FUNCTION_BLOCK LevelSensors (* Composite Function Block Type *)
  (* Standard: 61499-2 *)
  (* Version 0.0, 6/20/2016, Andrei, nxtControl GmbH, template *)
  PACKAGE Main;
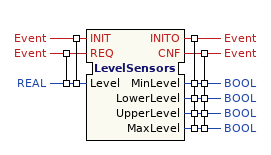
  EVENT_INPUT
    INIT WITH Level; (* Initialization Request *)
    REQ WITH Level; (* Normal Execution Request *)
  END_EVENT
  EVENT_OUTPUT
    INITO WITH MinLevel, LowerLevel, UpperLevel, MaxLevel; (* Initialization Confirm *)
    CNF WITH MinLevel, LowerLevel, UpperLevel, MaxLevel; (* Execution Confirmation *)
  END_EVENT
  VAR_INPUT
    Level : REAL; (* Input event qualifier *)
  END_VAR
  VAR_OUTPUT
    MinLevel : BOOL; (* Output event qualifier *)
    LowerLevel : BOOL;
    UpperLevel : BOOL;
    MaxLevel : BOOL;
  END_VAR
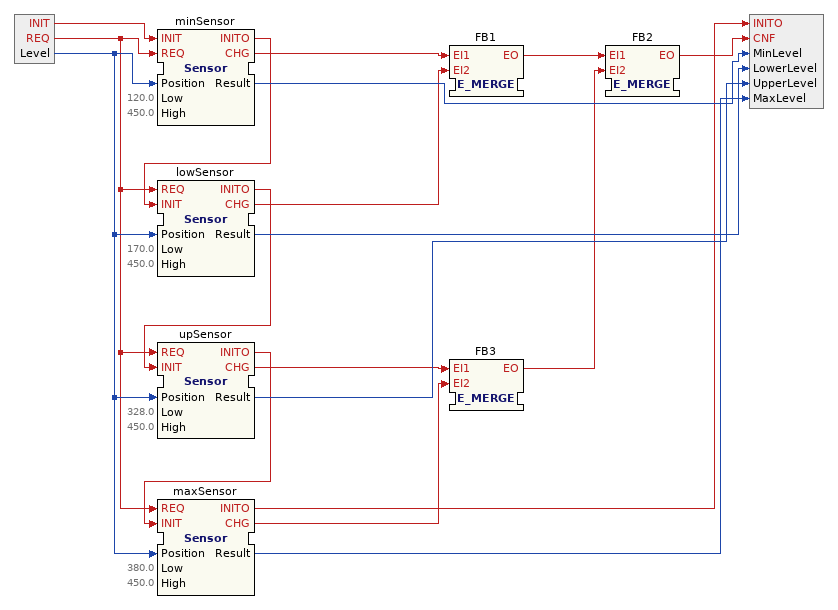
  FBS
    FB1 : E_MERGE;
    FB2 : E_MERGE;
    FB3 : E_MERGE;
    minSensor : Sensor(Low := 120.0, High := 450.0);
    lowSensor : Sensor(Low := 170.0, High := 450.0);
    upSensor : Sensor(Low := 328.0, High := 450.0);
    maxSensor : Sensor(Low := 380.0, High := 450.0);
  END_FBS
  EVENT_CONNECTIONS
    INIT TO minSensor.INIT;
    REQ TO minSensor.REQ;
    REQ TO lowSensor.REQ;
    REQ TO upSensor.REQ;
    REQ TO maxSensor.REQ;
    minSensor.INITO TO lowSensor.INIT;
    lowSensor.INITO TO upSensor.INIT;
    upSensor.INITO TO maxSensor.INIT;
    maxSensor.INITO TO INITO;
    FB1.EO TO FB2.EI1;
    FB3.EO TO FB2.EI2;
    FB2.EO TO CNF;
    minSensor.CHG TO FB1.EI1;
    upSensor.CHG TO FB3.EI1;
    maxSensor.CHG TO FB3.EI2;
    lowSensor.CHG TO FB1.EI2;
  END_CONNECTIONS
  DATA_CONNECTIONS
    Level TO minSensor.Position;
    Level TO lowSensor.Position;
    Level TO upSensor.Position;
    Level TO maxSensor.Position;
    minSensor.Result TO MinLevel;
    lowSensor.Result TO LowerLevel;
    upSensor.Result TO UpperLevel;
    maxSensor.Result TO MaxLevel;
  END_CONNECTIONS
END_FUNCTION_BLOCK
